(*
SPDX-FileCopyrightText: © 2026 Oleksandr Tiutyk <trofimich@gmail.com>
SPDX-License-Identifier: MIT
License: https://opensource.org/license/mit
*)

(*!
<summary>Common base interface for workflow activities and conditions participating in a workflow hierarchy.</summary>
<description>
The standard construction APIs enforce one borrowed parent slot per instance, acyclic parent links and
fixed workflow association. Unassociated subtrees may inherit an owner after attachment; associated children
require an already associated parent with the same owner. Configuration requires PASSIVE_READY throughout
the parent chain and owning workflow. Callers keep the tree live and stable, use one task, avoid reentry
and do not copy ownership-bearing instances by value. These rules do not provide cross-task synchronization.
</description>
*)

INTERFACE IWorkflowElement EXTENDS IVariableLookup, TOF_Core.INamed

(*!
<summary>Returns the parent workflow element in the hierarchy, or 0 for a root element.</summary>
*)
{attribute 'monitoring' := 'call'}
PROPERTY Parent : IWorkflowElement
GET
END_GET
END_PROPERTY

(*!
<summary>Returns the workflow that hosts this element, or 0 when not associated with a workflow.</summary>
*)
{attribute 'monitoring' := 'call'}
PROPERTY Workflow : IWorkflow
GET
END_GET
END_PROPERTY

END_INTERFACE

(* stored: Version 1.1.0.1
   Itf IWorkflowElement: Id {9f2cf0e1-485a-4f9c-a99d-72fe864dad44}
   Property Parent: Id {cfa98d13-c681-4820-8998-f8a3411bc85d}
   Get Get: Id {7ec43eb9-38c8-4405-b62f-59911e7d0170}
   Property Workflow: Id {1d31faa1-77cb-4600-b9ac-1ebaa9abd2ff}
   Get Get: Id {7fde95c5-a31e-46bf-a4f2-cad5094ce479} *)
